// Nature d'une position planaire (docs/05 § 6.1)
{attribute 'qualified_only'}
{attribute 'strict'}
TYPE E_PlanarPosKind :
(
    Work := 0,
    Queue := 1,
    Buffer := 2,
    Park := 3
) USINT;
END_TYPE

(* stored: Version 1.1.0.1, ProductVersion 3.1.4024.12
   DUT E_PlanarPosKind: Id {e7dcbfdc-efda-5d0f-b278-cfe02e5d063d} *)
